(* PLC project zarechnaya.project, CODESYS CODESYS V3.5 SP17 Patch 3 *)
(* stored: creationDateTime 2026-10-20T05:42:22.2931425, modificationDateTime 1601-01-01T03:00:00 *)

(* PRG_Backwash — промывка фильтра (SFC, PROGRAM: таймауты, N/S/R/P). Шаги: Idle (начальный) → [xStart] → Drain → [Drain.t >= T#2S] → Wash → [Wash.t >= T#3S] → Rinse → [Rinse.t >= T#1S OR xAbort] → Idle. Действия (IEC): Drain — N ActDrain (iDrainTicks += 1), S ActValve (iValveTicks += 1); Wash — N ActWash (iWashTicks += 1), P ActCount (iCycles += 1); Rinse — R ActValve, N ActRinse (iRinseTicks += 1). Порядок цикла — справка CODESYS (lower/sfc.py); IEC-действие исполняется ещё раз после деактивации (последний вызов с Q = FALSE). entry/exit-действия в CODESYS 3.5.17 не импортируются из PLCopen (M0: N), поэтому в кейсе их нет — автомат c2s7 их поддерживает (unit-тесты). *)
PROGRAM PRG_Backwash
  VAR_INPUT
    xStart : BOOL;
    xAbort : BOOL;
  END_VAR
  VAR_OUTPUT
    iDrainTicks : INT;
    iValveTicks : INT;
    iWashTicks : INT;
    iCycles : INT;
    iRinseTicks : INT;
  END_VAR

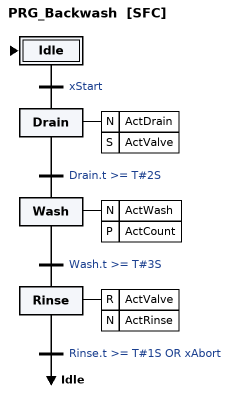
INITIAL_STEP Idle:
END_STEP
TRANSITION FROM Idle TO Drain
  := xStart;
END_TRANSITION
STEP Drain:
  ActDrain(N);
  ActValve(S);
END_STEP
TRANSITION FROM Drain TO Wash
  := Drain.t >= T#2S;
END_TRANSITION
STEP Wash:
  ActWash(N);
  ActCount(P);
END_STEP
TRANSITION FROM Wash TO Rinse
  := Wash.t >= T#3S;
END_TRANSITION
STEP Rinse:
  ActValve(R);
  ActRinse(N);
END_STEP
TRANSITION FROM Rinse TO Idle
  := Rinse.t >= T#1S OR xAbort;
END_TRANSITION

ACTION ActDrain:
                iDrainTicks := iDrainTicks + 1;

              
END_ACTION

ACTION ActValve:
                iValveTicks := iValveTicks + 1;

              
END_ACTION

ACTION ActWash:
                iWashTicks := iWashTicks + 1;

              
END_ACTION

ACTION ActCount:
                iCycles := iCycles + 1;

              
END_ACTION

ACTION ActRinse:
                iRinseTicks := iRinseTicks + 1;

              
END_ACTION
END_PROGRAM
